FUNCTION_BLOCK ABSTRACT FB_AnyValue IMPLEMENTS I_OtlpValue

(*
	Releases this value and clears the caller's pointer to it: call it as p^.delete(pSelf:=p).
	pSelf is cleared before the value is freed, so the caller never keeps a dangling pointer.
	A pointer to any other object is refused and left untouched, and nothing is released.
*)
METHOD ABSTRACT delete : BOOL
VAR_IN_OUT
	pSelf: POINTER TO FB_AnyValue;
END_VAR
END_METHOD

PROPERTY ABSTRACT eType : E_ValueType
GET
END_GET
END_PROPERTY

(* deallocates all data owned by the value without deleting the object itself.*)
METHOD ABSTRACT free
END_METHOD

END_FUNCTION_BLOCK

(* stored: Version 1.1.0.1
   POU FB_AnyValue: Id {ded18306-68d2-4405-b771-761d4aa3f677}, SpecialFunc None
   Method delete: Id {86d3a7ce-6868-4d24-99f2-1892df9a286c}
   Property eType: Id {516a8d71-2631-45bf-9dd6-2becf5f4e651}
   Get Get: Id {7b0372bd-bf22-4369-8533-5ee73c5848f0}
   Method free: Id {7cccd8b3-2131-4b23-8124-c1d537a212e8} *)
